// Parametri macchina scritti dall'HMI (HMI -> PLC); diventano effettivi con il comando WriteParameters.
TYPE ST_HmiParam :
STRUCT
	bEnableSirenOverride	: BOOL;
	aAxis					: ARRAY[1..Core_Param.MAX_AXIS] OF ST_HmiAxisParam;
END_STRUCT
END_TYPE

(* stored: Version 1.1.0.1, ProductVersion 3.1.4024.12
   DUT ST_HmiParam: Id {57c1015d-2d4f-4ba0-918c-d81d5122d2d0} *)
